VISUALIZATION VisuNoMan  // 2x2
END_VISUALIZATION

(* stored: Version 1.1.0.1
   Visu VisuNoMan: Id {e845e8e7-c27e-4fb1-ac54-6a44a39bcef4} *)
